// TIA Portal V20 export
// export: Created 2026-10-11T05:31:07.8219902Z, ExportSetting WithDefaults, DisplayName Totally Integrated Automation Portal, DisplayVersion V20, DisplayName TIA Portal Openness, DisplayVersion V20, DisplayName TIA Portal Teamcenter Gateway, DisplayVersion V20, DisplayName TIA Portal Version Control Interface, DisplayVersion V20, DisplayName SINAMICS Startdrive Advanced, DisplayVersion V20 SP1 Update 2, DisplayName SINAMICS Startdrive G110M, G120, G120C, G120D, G120P, G115D, DisplayVersion V20 SP1 Update 2, DisplayName SINAMICS Startdrive G130, G150, S120, S150, SINAMICS MV, G220, S200, S210, DisplayVersion V20 SP1 Update 2, DisplayName STEP 7 Professional, DisplayVersion V20, DisplayName STEP 7 Safety, DisplayVersion V20, DisplayName WinCC Basic/Comfort/Advanced, DisplayVersion V20, DisplayName WinCC Professional, DisplayVersion V20, DisplayName WinCC Unified, DisplayVersion V20
FUNCTION "FRK_Fault" : Void   // FC8, SCL
{ S7_Optimized_Access := 'TRUE' }
VERSION : 0.1
// stored: AutoNumber true, IsIECCheckEnabled false, SetENOAutomatically false, UDAEnableTagReadback false
   VAR_INPUT
      ReasonCode : DInt;
      Description : WString;
   END_VAR
   VAR_IN_OUT
      Core : "FRK_Core";
      Status : "ST_ModuleStatus";
   END_VAR
BEGIN

   IF #Core.Exec = 3 THEN
       RETURN;
   END_IF;
   "FRK_Diagnostic"(Status := #Status,
                    ReasonCode := #ReasonCode,
                    Description := #Description,
                    Severity := 1);
   "FRK_Rationalize"(Diag := #Status.Diagnostic);
   #Core.Exec := 3;
   #Core.Step := 0;
   #Core.Dispatch := FALSE;
   #Core.DiagTouched := TRUE;
END_FUNCTION
